(* IEC 61131-3 sources: Test-Git_ESME26/TestProgettoESME_26.fbsproj/PacDriveLib Migration/Motion/Homing/PDL_FB_SetDrvEncPos.fb.st^, 4 files *)

(* ---- diResultSetDrvEncPos.prop.st ---- *)
PROPERTY PUBLIC diResultSetDrvEncPos : DINT
__GETTERDECLARATION__
VAR
END_VAR
__GETTERIMPLEMENTATION__
diResultSetDrvEncPos := diResultSetDrvEnc_loc;

(* ---- ifDeviceType.prop.st ---- *)
PROPERTY PUBLIC ifDeviceType : DeviceTypeInterfaces.IF_Device_Type
__SETTERDECLARATION__
VAR
END_VAR
__SETTERIMPLEMENTATION__
ifDeviceType_loc := ifDeviceType;

(* ---- lrPosition.prop.st ---- *)
PROPERTY PUBLIC lrPosition : LREAL
__SETTERDECLARATION__
VAR
END_VAR
__SETTERIMPLEMENTATION__
lrPosition_loc := lrPosition;

(* ---- xDone.prop.st ---- *)
PROPERTY xDone : BOOL
__SETTERDECLARATION__
VAR
END_VAR
__SETTERIMPLEMENTATION__
xDone_loc := xDone;
__GETTERDECLARATION__
VAR
END_VAR
__GETTERIMPLEMENTATION__
xDone := xDone_loc;
